Staubli VAL3: io.dtx


